__TRY
	_Loaded := _LoadLoader.Load(
		reader := _LoadReader,
		root := _LoadReader.Parse(document := _ConfigDocument),
		factory := THIS^,
		dependencyFactory := THIS^,
		resolver := THIS^,
		binder := THIS^
	);
__CATCH(exceptionCode)
	exception := TOF_Core.ExceptionManager.GetLastException(
		exceptionCode := exceptionCode,
		catchPointNamespaceName := NamespaceName,
		catchPointPOUName := __POUNAME(),
		catchPointPosition := __POSITION()
	);
	caught := exception <> 0 AND_THEN __QUERYINTERFACE(exception, configurationError);
__ENDTRY

IF NOT caught AND_THEN exception <> 0 THEN
	assertions.ThatBool(
		actual := FALSE,
		message := TO_WSTRING(TOF_Core.Strings.Concat255('Unbound workflow load: ', TO_STRING(exception.GetMessage())))
	).IsTrue();
ELSE
	assertions.ThatBool(
		actual := caught AND_THEN _Loaded = 0,
		message := "Unresolved required PLC variable must abort and roll back load"
	).IsTrue();
END_IF

IF _Loaded <> 0 THEN
	assertions.ThatBool(
		actual := TryReleaseLoadedWorkflow(),
		message := "Release any unexpected workflow after the unbound load"
	).IsTrue();
END_IF

TOF_Core.DynamicMemoryManager.RaiseIfAllocationFailed();

_BindLoadVariables := TRUE;
_LoadExternal := 11;
caught := FALSE;
__TRY
	_Loaded := _LoadLoader.Load(
		reader := _LoadReader,
		root := _LoadReader.Parse(document := _ConfigDocument),
		factory := THIS^,
		dependencyFactory := THIS^,
		resolver := THIS^,
		binder := THIS^
	);
__CATCH(exceptionCode)
	caught := TRUE;
	exception := TOF_Core.ExceptionManager.GetLastException(
		exceptionCode := exceptionCode,
		catchPointNamespaceName := NamespaceName,
		catchPointPOUName := __POUNAME(),
		catchPointPosition := __POSITION()
	);

	IF exception <> 0 THEN
		assertions.ThatBool(
			actual := FALSE,
			message := TO_WSTRING(TOF_Core.Strings.Concat255('Bound workflow load: ', TO_STRING(exception.GetMessage())))
		).IsTrue();
	ELSE
		assertions.ThatBool(
			actual := FALSE,
			message := TO_WSTRING(TOF_Core.Strings.Concat255('Bound workflow load raised PLC exception ', TO_STRING(exceptionCode)))
		).IsTrue();
	END_IF
__ENDTRY

IF NOT caught THEN
	assertions.ThatBool(
		actual := _Loaded <> 0 AND_THEN _Loaded.State = TOF_Workflow.WORKFLOW_ELEMENT_STATE.PASSIVE_READY,
		message := "Loaded workflow must be ready without auto-starting"
	).IsTrue();
END_IF

IF _Loaded <> 0 THEN
	_Loaded.RequestStart();

	FOR i := 1 TO 6 DO
		IF _Loaded.Busy THEN
			_Loaded.Execute();
		END_IF
	END_FOR

	assertions.ThatBool(
		actual := _Loaded.State = TOF_Workflow.WORKFLOW_ELEMENT_STATE.PASSIVE_COMPLETED,
		message := "Loaded workflow must execute embedded and external tasks and branch assignment"
	).IsTrue();

	ready := __QUERYINTERFACE(_Loaded.RootActivity, ifElse)
		AND_THEN __QUERYINTERFACE(_Loaded.RootActivity, rootScope)
		AND_THEN __QUERYINTERFACE(ifElse.Condition, conditionScope);
	assertions.ThatBool(
		actual := ready,
		message := "Loaded root and condition must expose declaration containers"
	).IsTrue();

	IF ready THEN
		localStep := rootScope.GetDeclaredElement(name := 'LocalStep', index := 0);
		limitElement := rootScope.GetDeclaredElement(name := 'Limits', index := 1);
		thresholdElement := conditionScope.GetDeclaredElement(name := 'Threshold', index := 0);
		assertions.ThatBool(
			actual := localStep.AsUInt() = 11 AND_THEN limitElement.AsUInt() = 8 AND_THEN thresholdElement.AsUInt() = 3,
			message := "Loaded execution must update target declaration and preserve array and condition values"
		).IsTrue();

		limitElement.ChangeValueByAny(value := mutated);
		thresholdElement.ChangeValueByAny(value := mutated);
		_Loaded.RequestReset();

		assertions.ThatBool(
			actual := _Loaded.State = TOF_Workflow.WORKFLOW_ELEMENT_STATE.PASSIVE_READY
				AND_THEN localStep.AsUInt() = 3
				AND_THEN limitElement.AsUInt() = 8
				AND_THEN thresholdElement.AsUInt() = 3,
			message := "Resetting a loaded workflow must restore activity and condition declarations in place"
		).IsTrue();
	END_IF

	assertions.ThatBool(
		actual := TryReleaseLoadedWorkflow(),
		message := "Release the dynamically loaded workflow"
	).IsTrue();
END_IF

_LoadSource.DisposeDynamicChildren();
TOF_Core.DynamicMemoryManager.RaiseIfAllocationFailed();
END_METHOD

(*!
<summary>Verifies that workflow element deserialization rejects null context and context-free succeeds.</summary>
<description>
A workflow element requiring a loader raises WorkflowConfiguration when deserialized with context = 0.
A context-free element (DelayActivity) succeeds when deserialized with context = 0.
</description>
<param name="assertions">Valid assertion context borrowed from the active case.</param>
*)
METHOD PRIVATE testDeserializeNullContextRejection
VAR_INPUT
	assertions : REFERENCE TO TOF_Testing.Assertions;
END_VAR
VAR
	workflowNode : TOF_Core.CONFIGURATION_NODE;
	delayNode : TOF_Core.CONFIGURATION_NODE;
	caught : BOOL;
	exceptionCode : __SYSTEM.ExceptionCode;
	exception : TOF_Core.IException;
	configurationError : TOF_Workflow.IWorkflowConfigurationException;
END_VAR
_ConfigWriter.Serialize(source := _NullContextSequence, document := _ConfigDocument);
workflowNode := _LoadReader.Parse(document := _ConfigDocument);

caught := FALSE;
__TRY
	_NullContextSequence.Deserialize(reader := _LoadReader, node := workflowNode, context := 0);
__CATCH(exceptionCode)
	exception := TOF_Core.ExceptionManager.GetLastException(
		exceptionCode := exceptionCode,
		catchPointNamespaceName := NamespaceName,
		catchPointPOUName := __POUNAME(),
		catchPointPosition := __POSITION()
	);
	caught := __QUERYINTERFACE(exception, configurationError);
__ENDTRY

assertions.ThatBool(
	actual := caught,
	message := "Workflow element requiring loader must reject null deserialization context"
).IsTrue();

_NullContextDelay.Interval := T#5S;
_ConfigWriter.Serialize(source := _NullContextDelay, document := _ConfigDocument);
delayNode := _LoadReader.Parse(document := _ConfigDocument);

caught := FALSE;
__TRY
	_NullContextDelay.Deserialize(reader := _LoadReader, node := delayNode, context := 0);
__CATCH(exceptionCode)
	caught := TRUE;
__ENDTRY

assertions.ThatBool(
	actual := caught,
	message := "Context-free workflow element must succeed with null deserialization context"
).IsFalse();
assertions.ThatTime(
	actual := _NullContextDelay.Interval,
	message := "Delay interval must be restored"
).ToBe(expected := T#5S);

TOF_Core.DynamicMemoryManager.RaiseIfAllocationFailed();
END_METHOD

(*!
<summary>Verifies formatting and parsing of logical and comparison operators.</summary>
<param name="assertions">Valid assertion context borrowed from the active case.</param>
*)
METHOD PRIVATE testOperatorSerialization
VAR_INPUT
	assertions : REFERENCE TO TOF_Testing.Assertions;
END_VAR
VAR
	caught : BOOL;
	exceptionCode : __SYSTEM.ExceptionCode;
	exception : TOF_Core.IException;
	configurationError : TOF_Workflow.IWorkflowConfigurationException;
	parsedComp : TOF_Workflow.COMPARISON_OPERATOR;
	parsedLog : TOF_Workflow.LOGICAL_OPERATOR;
END_VAR
// Format comparison operators
assertions.ThatString(
	actual := TOF_Workflow.Workflows.FormatComparisonOperator(comparisonOperator := TOF_Workflow.COMPARISON_OPERATOR.EQUAL),
	message := "Format EQUAL"
).ToBe(expected := '=');
assertions.ThatString(
	actual := TOF_Workflow.Workflows.FormatComparisonOperator(comparisonOperator := TOF_Workflow.COMPARISON_OPERATOR.NOT_EQUAL),
	message := "Format NOT_EQUAL"
).ToBe(expected := '<>');
assertions.ThatString(
	actual := TOF_Workflow.Workflows.FormatComparisonOperator(comparisonOperator := TOF_Workflow.COMPARISON_OPERATOR.LESS_THAN),
	message := "Format LESS_THAN"
).ToBe(expected := '<');
assertions.ThatString(
	actual := TOF_Workflow.Workflows.FormatComparisonOperator(comparisonOperator := TOF_Workflow.COMPARISON_OPERATOR.LESS_THAN_OR_EQUAL),
	message := "Format LESS_THAN_OR_EQUAL"
).ToBe(expected := '<=');
assertions.ThatString(
	actual := TOF_Workflow.Workflows.FormatComparisonOperator(comparisonOperator := TOF_Workflow.COMPARISON_OPERATOR.GREATER_THAN),
	message := "Format GREATER_THAN"
).ToBe(expected := '>');
assertions.ThatString(
	actual := TOF_Workflow.Workflows.FormatComparisonOperator(comparisonOperator := TOF_Workflow.COMPARISON_OPERATOR.GREATER_THAN_OR_EQUAL),
	message := "Format GREATER_THAN_OR_EQUAL"
).ToBe(expected := '>=');

// Parse comparison operators and synonyms
parsedComp := TOF_Workflow.Workflows.ParseComparisonOperator(rawOperator := '=');
assertions.ThatBool(actual := parsedComp = TOF_Workflow.COMPARISON_OPERATOR.EQUAL, message := "Parse =").IsTrue();

parsedComp := TOF_Workflow.Workflows.ParseComparisonOperator(rawOperator := '==');
assertions.ThatBool(actual := parsedComp = TOF_Workflow.COMPARISON_OPERATOR.EQUAL, message := "Parse ==").IsTrue();

parsedComp := TOF_Workflow.Workflows.ParseComparisonOperator(rawOperator := '<>');
assertions.ThatBool(
	actual := parsedComp = TOF_Workflow.COMPARISON_OPERATOR.NOT_EQUAL,
	message := "Parse <>"
).IsTrue();

parsedComp := TOF_Workflow.Workflows.ParseComparisonOperator(rawOperator := '!=');
assertions.ThatBool(
	actual := parsedComp = TOF_Workflow.COMPARISON_OPERATOR.NOT_EQUAL,
	message := "Parse !="
).IsTrue();

parsedComp := TOF_Workflow.Workflows.ParseComparisonOperator(rawOperator := '<');
assertions.ThatBool(
	actual := parsedComp = TOF_Workflow.COMPARISON_OPERATOR.LESS_THAN,
	message := "Parse <"
).IsTrue();

parsedComp := TOF_Workflow.Workflows.ParseComparisonOperator(rawOperator := '<=');
assertions.ThatBool(
	actual := parsedComp = TOF_Workflow.COMPARISON_OPERATOR.LESS_THAN_OR_EQUAL,
	message := "Parse <="
).IsTrue();

parsedComp := TOF_Workflow.Workflows.ParseComparisonOperator(rawOperator := '>');
assertions.ThatBool(
	actual := parsedComp = TOF_Workflow.COMPARISON_OPERATOR.GREATER_THAN,
	message := "Parse >"
).IsTrue();

parsedComp := TOF_Workflow.Workflows.ParseComparisonOperator(rawOperator := '>=');
assertions.ThatBool(
	actual := parsedComp = TOF_Workflow.COMPARISON_OPERATOR.GREATER_THAN_OR_EQUAL,
	message := "Parse >="
).IsTrue();

// Invalid comparison operator
caught := FALSE;
__TRY
	parsedComp := TOF_Workflow.Workflows.ParseComparisonOperator(rawOperator := 'INVALID');
__CATCH(exceptionCode)
	exception := TOF_Core.ExceptionManager.GetLastException(
		exceptionCode := exceptionCode,
		catchPointNamespaceName := NamespaceName,
		catchPointPOUName := __POUNAME(),
		catchPointPosition := __POSITION()
	);
	caught := __QUERYINTERFACE(exception, configurationError);
__ENDTRY
assertions.ThatBool(actual := caught, message := "Unknown comparison operator must raise").IsTrue();

// Format logical operators
assertions.ThatString(
	actual := TOF_Workflow.Workflows.FormatLogicalOperator(logicalOperator := TOF_Workflow.LOGICAL_OPERATOR.AND_),
	message := "Format AND_"
).ToBe(expected := 'AND');
assertions.ThatString(
	actual := TOF_Workflow.Workflows.FormatLogicalOperator(logicalOperator := TOF_Workflow.LOGICAL_OPERATOR.OR_),
	message := "Format OR_"
).ToBe(expected := 'OR');

// Parse logical operators
parsedLog := TOF_Workflow.Workflows.ParseLogicalOperator(rawOperator := 'AND');
assertions.ThatBool(actual := parsedLog = TOF_Workflow.LOGICAL_OPERATOR.AND_, message := "Parse AND").IsTrue();

parsedLog := TOF_Workflow.Workflows.ParseLogicalOperator(rawOperator := 'and');
assertions.ThatBool(
	actual := parsedLog = TOF_Workflow.LOGICAL_OPERATOR.AND_,
	message := "Parse and lowercase"
).IsTrue();

parsedLog := TOF_Workflow.Workflows.ParseLogicalOperator(rawOperator := 'AND_');
assertions.ThatBool(actual := parsedLog = TOF_Workflow.LOGICAL_OPERATOR.AND_, message := "Parse AND_").IsTrue();

parsedLog := TOF_Workflow.Workflows.ParseLogicalOperator(rawOperator := 'OR');
assertions.ThatBool(actual := parsedLog = TOF_Workflow.LOGICAL_OPERATOR.OR_, message := "Parse OR").IsTrue();

parsedLog := TOF_Workflow.Workflows.ParseLogicalOperator(rawOperator := 'or');
assertions.ThatBool(
	actual := parsedLog = TOF_Workflow.LOGICAL_OPERATOR.OR_,
	message := "Parse or lowercase"
).IsTrue();

parsedLog := TOF_Workflow.Workflows.ParseLogicalOperator(rawOperator := 'OR_');
assertions.ThatBool(actual := parsedLog = TOF_Workflow.LOGICAL_OPERATOR.OR_, message := "Parse OR_").IsTrue();

// Invalid logical operator
caught := FALSE;
__TRY
	parsedLog := TOF_Workflow.Workflows.ParseLogicalOperator(rawOperator := 'XOR');
__CATCH(exceptionCode)
	exception := TOF_Core.ExceptionManager.GetLastException(
		exceptionCode := exceptionCode,
		catchPointNamespaceName := NamespaceName,
		catchPointPOUName := __POUNAME(),
		catchPointPosition := __POSITION()
	);
	caught := __QUERYINTERFACE(exception, configurationError);
__ENDTRY
assertions.ThatBool(actual := caught, message := "Unknown logical operator must raise").IsTrue();

TOF_Core.DynamicMemoryManager.RaiseIfAllocationFailed();
END_METHOD

(*!
<summary>Attempts to release the owned result of a configuration load.</summary>
<description>Clears the stored alias before release. Succeeds if no workflow is owned.</description>
*)
METHOD TryReleaseLoadedWorkflow : BOOL
VAR
	instance : TOF_Core.IObject;
END_VAR
IF _Loaded = 0 THEN
	TryReleaseLoadedWorkflow := TRUE;

	RETURN;
END_IF

instance := _Loaded;
_Loaded := 0;
TryReleaseLoadedWorkflow := TOF_Core.Memory.TryReleaseDynamicObject(instance := instance);
END_METHOD

(*!
<summary>Clears a still-owned loaded workflow if the fixture is unloaded before case teardown.</summary>
<param name="bInCopyCode">TwinCAT copy-code exit marker. Leave copied ownership with the new instance.</param>
*)
METHOD FB_exit : BOOL
VAR_INPUT
	bInCopyCode : BOOL;
END_VAR
IF NOT bInCopyCode THEN
	TryReleaseLoadedWorkflow();
END_IF

FB_exit := TRUE;
END_METHOD

END_FUNCTION_BLOCK

(* stored: Version 1.1.0.1
   POU WorkflowContractTestFixture: Id {c420144d-dae1-4264-b0c8-03a582be053e}, SpecialFunc None
   Method ExecuteScenario: Id {6d02c419-d0c8-45cb-b367-0551d8d0f84d}
   Property ClassName: Id {96eb901b-f5de-49b0-bbcc-736ee2909b9b}
   Get Get: Id {682bf6bf-f8f2-4590-88ad-869259d5bca2}
   Property NamespaceName: Id {00ea1253-3cad-4942-9392-0a19c1354af1}
   Get Get: Id {256f3a94-281b-458b-bc8f-49bec55ef2d4}
   Property SelfSize: Id {7b82c98b-a45d-412e-82b9-f5d724c741d7}
   Get Get: Id {29ae5c68-f508-4929-afab-5a9b493616ac}
   Method testBoundaryDiagnostics: Id {adf9b6f6-08b7-404f-977b-06b3d4d5a22c}
   Method testCatchCleanupBoundary: Id {15577c12-1b83-427f-a3c6-edb36a3b31ec}
   Method testConcreteMetadata: Id {19af6d1d-6adf-419a-abf8-378e1113f396}
   Method testConditionScopePrecedence: Id {d54cfd66-8e51-4e3b-8ef1-bcd56fa4e3ee}
   Method testConditionTopology: Id {b1cbcc93-94b7-4d1f-aa83-86cf97d1f3c5}
   Method testDelayLifecycle: Id {8a705608-0fe1-495e-a6d9-5e201d173db0}
   Method testInitializationRetry: Id {63f3bffc-b980-4de2-827d-f9b07c8a03d3}
   Method testInvokeConfiguration: Id {c00f8cc8-9765-4529-9eb8-6aaa22393e11}
   Method testParentSetters: Id {372e3208-2548-408e-85ab-4efe636a6d24}
   Method testRootAssociation: Id {114a78e6-e29d-4e2f-9898-e5660c5c4f60}
   Method testSequenceTopology: Id {dd172252-0707-47a8-b182-7f7e89931c3a}
   Method testTaskAbortDuringSuspend: Id {51cb9f83-b866-4ad0-b866-bd3c07c2169b}
   Method testTaskCompletionDuringSuspend: Id {61c087d0-ad3f-4074-9944-38a066a82671}
   Method testTaskFailureDuringSuspend: Id {d4e3be94-3fa0-40cf-a203-fe128a3485be}
   Method testTaskReleaseFailureDuringCancel: Id {d8bd19e1-fb81-4153-aa67-873b0badd418}
   Method testVariableLookup: Id {a0945ab8-8ea1-4142-a5cf-84119b851dfb}
   Method testWorkflowIsolation: Id {b23d391b-b15f-4c8c-97eb-27107f3a5ab5}
   Method testDeclaredVariableReset: Id {88fce0b7-1178-4ac8-8f15-1fcf2375221d}
   Method testDeclaredVariableValidation: Id {e7938411-1f9d-427d-b002-9a332b8ba8f1}
   Method testTransitionDiagnostics: Id {fbcb0ede-daec-44f8-b076-0b6e0b28e502}
   Method CreateElement: Id {b350a52f-ef28-4138-84f4-fe6c914ab79a}
   Method testFactoryDeclarations: Id {96c2d6be-c9ed-4710-b132-79636718eda7}
   Method testArrayValidation: Id {c0b67d55-8aff-4a4a-b740-76f409bc9946}
   Method testWriteConfiguration: Id {c20c2bfa-8c1e-4a82-a125-8f08bdad54b0}
   Method testDependencyBindings: Id {4f68a902-c396-448e-8518-ecdb48a31599}
   Method CreateDependency: Id {e8bcc63f-b77a-44fc-a5cf-2712acf9b5ce}
   Method ResolveExternal: Id {486c7ba3-eb9c-4d1e-90f9-49250a5b16d2}
   Method BindVariables: Id {2256e760-cfa4-4f34-be80-fcd785ebbc1e}
   Method testLoadConfiguration: Id {846b9dc0-e206-4ab5-b87c-42169368526e}
   Method testDeserializeNullContextRejection: Id {f28d6d68-5863-49f9-9dc3-cdffc37a855f}
   Method testOperatorSerialization: Id {76631bbb-6383-45e4-a2fc-c6d60459c699}
   Method TryReleaseLoadedWorkflow: Id {e3970f7b-166e-4eae-afff-a7fa7068e7d1}
   Method FB_exit: Id {b63d2f44-d576-41b8-abef-9c96db90411b} *)
